PROGRAM PRG_CNCDiagnostics
VAR
	fbCNCDiagnosisUpload : FB_CNCDiagnosisUpload;
	bUploadDiagData: BOOL;
END_VAR

fbCNCDiagnosisUpload(
	bExecute:= bUploadDiagData, 
	strFileName:= 'C:\temp\diag_data.txt', 
	nHistory:= 0, 
	strTopic:= 'ALL', 
	bBusy=> , 
	bError=> , 
	nErrorID=> );

END_PROGRAM

(* stored: Version 1.1.0.1
   POU PRG_CNCDiagnostics: Id {6696336b-5503-4742-bdb3-3e9cfb3c1521}, SpecialFunc None *)
